// Forçage d'un mover (docs/12 § 4)
{attribute 'pack_mode' := '1'}
TYPE ST_MoverForce :
STRUCT
    bOutOfService : BOOL;
    bImmediate : BOOL;
    nReason : USINT;
    tSince : LINT;
    sBy : STRING(24);
END_STRUCT
END_TYPE

(* stored: Version 1.1.0.1, ProductVersion 3.1.4024.12
   DUT ST_MoverForce: Id {a0c106d9-f43e-568b-95b8-6e5eddd978bc} *)
